(* IEC 61131-3 sources: 2026_Projet_YGO_ExcavatriceDragage/CODE_BACKUP/CODE_20260803_avant_ee4d08b/ACQUISITION, 1 file *)

(* ---- FB_AcquisitionLegacyBridge.st ---- *)
(* ═══════════════════════════════════════════════════════════════
   📡 FB_AcquisitionLegacyBridge — Pont temporaire acquisition historique
   ───────────────────────────────────────────────────────────────
   📄 Docs : DOC/AF_Partie-06_Acquisition_Qualification_IO_v2.0.md §2 ;
            DOC/AF_Partie-13_Fonction_Simulation_v2.0.md
   ⚙️ Pont ST temporaire appelé exclusivement par PRG_02_Acquisition_CFC.xml.
   🎯 Rôle unique : produire l'image matérielle HwIn consommée par le reste
      du programme. Aucune décision métier (SafeStop, mode, commande) ici.
   🔗 Producteur unique de HwIn ; consommateurs = PRG_01_Inputs_LD et suivants.
   ═══════════════════════════════════════════════════════════════ *)

FUNCTION_BLOCK FB_AcquisitionLegacyBridge

VAR_OUTPUT
    HwReal                   : ST_HardwareImage;  (* Image matérielle brute lue sur le terrain *)
    HwSim                    : ST_HardwareImage;  (* Image produite par le banc de simulation *)
    HwIn                     : ST_HardwareImage;  (* Image aiguillée réel/simulé *)
    WinchInputSourceChanged  : BOOL;              (* Pulse 1 cycle sur bascule réel/simulé domaine Winch *)

    // 🆕 Migration PRG_00_Inputs : positions Translation M3 exposées en sortie de programme
    TranslationPosTremie      : BOOL;   (* TRUE = translation en position Trémie *)
    TranslationPosPV          : BOOL;   (* TRUE = translation en zone pré-ralentissement PV *)
    TranslationPosP2          : BOOL;   (* TRUE = translation en position P2 *)
    TranslationPosP1          : BOOL;   (* TRUE = translation en position P1 *)
    TranslationPosMaintenance : BOOL;   (* TRUE = translation en position Maintenance *)

    // 🆕 Migration PRG_00_Inputs : retours variateur M3 filtrés (PT1 T#0MS = recopie legacy)
    M3_StatusWord_Filtered        : UINT;
    M3_ActualFrequencyHz_Filtered : UINT;

    // 🔗 Contrat public : anciennement lus à travers instPosDecoderM3.
    //    Les sorties rendent la migration XML transparente aux consommateurs.
    M3_LimitSwitchFwd          : BOOL;
    M3_LimitSwitchRev          : BOOL;
    M3_SensorWordIncoherent    : BOOL;
    M3_SensorsWord             : BYTE;
END_VAR

VAR
    (* ── Instances de traitement complexes ── *)
    instSimBench             : FB_SimBench;
    instJoystick             : FB_Joystick;
    instEncoderAbsM1         : FB_Encoder_Abs;
    instEncoderScaleM1       : FB_Encoder_Scale;
    instHomingM1             : FB_Encoder_Homing;
    instEncoderAbsM2         : FB_Encoder_Abs;
    instEncoderScaleM2       : FB_Encoder_Scale;
    instHomingM2             : FB_Encoder_Homing;
    instPosDecoderM3         : FB_Translation_PositionDecoder;

    (* ── Filtrage des retours variateur M3 (migration PRG_00_Inputs) ── *)
    instCycleTimeAcq            : FB_CycleTime;
    instFilterM3StatusWord      : FB_Filter_PT1;
    instFilterM3ActualFreqHz      : FB_Filter_PT1;

    (* ── Mémoire de la source Winch (front bascule réel/simulé) ── *)
    WinchInputSourceSimulated            : BOOL;
    PreviousWinchInputSourceSimulated    : BOOL;
    WinchInputSourceInitialized          : BOOL;
END_VAR

// === IMPLEMENTATION ===

// ─── §0 MATÉRIEL ──► HwReal (Acquisition brute unique) ─────────────────────────

// Winch M1 / M2 et codeurs
HwReal.Winch.M1_ContactorsReleased_DI := M1_ContactorsReleased_DI;
HwReal.Winch.M1_ThermalOk_DI          := M1_ThermalOk_DI;
HwReal.Winch.M1_BrakeIsOpen_DI        := M1_BrakeIsOpen_DI;

HwReal.Winch.M2_ContactorsReleased_DI := M2_ContactorsReleased_DI;
HwReal.Winch.M2_ThermalOk_DI          := M2_ThermalOk_DI;
HwReal.Winch.M2_BrakeIsOpen_DI        := M2_BrakeIsOpen_DI;

HwReal.Winch.M1M2_TopPositionFree_DI  := M1M2_TopPositionFree_DI;
HwReal.Winch.M2_TensionedCable_DI     := M2_TensionedCable_DI;

HwReal.Winch.COD1_PosValue            := COD1_PosValue;
HwReal.Winch.COD1_Alarms              := COD1_Alarms;
HwReal.Winch.COD1_Warnings            := COD1_Warnings;
HwReal.Winch.COD1_DeviceState         := COD1_CODEUR.GetDeviceState();

HwReal.Winch.COD2_PosValue            := COD2_PosValue;
HwReal.Winch.COD2_Alarms              := COD2_Alarms;
HwReal.Winch.COD2_Warnings            := COD2_Warnings;
HwReal.Winch.COD2_DeviceState         := COD2_CODEUR.GetDeviceState();

// Translation M3 et variateur AC600
HwReal.Translation.M3_PosTremie_DI      := M3_PosTremie_DI;
HwReal.Translation.M3_PosPV_DI          := M3_PosPV_DI;
HwReal.Translation.M3_PosP2_DI          := M3_PosP2_DI;
HwReal.Translation.M3_PosP1_DI          := M3_PosP1_DI;
HwReal.Translation.M3_PosMaintenance_DI := M3_PosMaintenance_DI;
HwReal.Translation.M3_BrakeIsOpen_DI    := M3_BrakeIsOpen_DI;
HwReal.Translation.M3_ThermalFeedback_DI:= M3_ThermalFeedback_DI; // 🆕 T96 — diagnostic seul (voie déjà mappée CODESYS, jamais lue jusqu'ici)
HwReal.Translation.M3_StatusWord        := M3_StatusWord;
HwReal.Translation.M3_ActualFrequencyHz := M3_ActualFrequencyHz;
HwReal.Translation.AC600_DeviceState    := AC600_ECAT_Drive.GetDeviceState();

// Opérateur / Joystick / bus CANopen
HwReal.Operator.JoyXRaw_ANA1      := JoyXRaw_ANA1;
HwReal.Operator.JoyYRaw_ANA2      := JoyYRaw_ANA2;
HwReal.Operator.JoyBtnRaw         := JoyBtnRaw;
HwReal.Operator.CanBusState       := CANbus.GetBusState();
HwReal.Operator.JOY1_DeviceState  := JOY1_JOYSTICK_MCB560_CO4201A.GetDeviceState();

// Sécurités / Communs Machine
HwReal.Machine.PowerContactorEngaged_DI   := PowerContactorEngaged_DI;
HwReal.Machine.EmergencyChainClosed_DI    := EmergencyChainClosed_DI;
HwReal.Machine.PhaseRotationOk_DI         := PhaseRotationOk_DI;
HwReal.Machine.BrakeThermalOk_DI          := BrakeThermalOk_DI;
HwReal.Machine.M1_M2_KoboldContactFond_DI := M1_M2_KoboldContactFond_DI;
HwReal.Machine.HydraulicThermalOk_DI      := HydraulicThermalOk_DI;

// ─── §0bis HwReal / SimBench ──► HwIn (Aiguillage simulation par domaine) ──────

instSimBench(
    Enable                   := GVL_Simulation.SimulationModeActive,
    M1_RelayFwd              := GVL_Global.M1RelayFwd,
    M1_RelayRev              := GVL_Global.M1RelayRev,
    M1_SpeedContactor_1      := GVL_Global.M1SpeedContactor1,
    M1_SpeedContactor_2      := GVL_Global.M1SpeedContactor2,
    M1_SpeedContactor_3      := GVL_Global.M1SpeedContactor3,
    M1_SpeedContactor_4      := GVL_Global.M1SpeedContactor4,
    M1_SpeedRefPct           := PRG_TREUILS_CFC.M1_SpeedRef_Active,
    M1_PresetTriggerCmd      := PRG_02_Encoders.instEncoderAbsM1.PresetTriggerCmd,
    M1_PresetValueOut        := PRG_02_Encoders.instEncoderAbsM1.PresetValueOut,
    M1_BrakeCmd              := GVL_Global.M1BrakeCmd,
    M2_RelayFwd              := GVL_Global.M2RelayFwd,
    M2_RelayRev              := GVL_Global.M2RelayRev,
    M2_SpeedContactor_1      := GVL_Global.M2SpeedContactor1,
    M2_SpeedContactor_2      := GVL_Global.M2SpeedContactor2,
    M2_SpeedContactor_3      := GVL_Global.M2SpeedContactor3,
    M2_SpeedContactor_4      := GVL_Global.M2SpeedContactor4,
    M2_SpeedRefPct           := PRG_TREUILS_CFC.M2_SpeedRef_Active,
    M2_PresetTriggerCmd      := PRG_02_Encoders.instEncoderAbsM2.PresetTriggerCmd,
    M2_PresetValueOut        := PRG_02_Encoders.instEncoderAbsM2.PresetValueOut,
    M2_BrakeCmd              := GVL_Global.M2BrakeCmd,
    M3_Direction             := PRG_TRANSLATION_CFC.M3_Direction_Active,
    M3_SpeedRefPct           := PRG_TRANSLATION_CFC.M3_SpeedRef_Active,
    M3_BrakeCmd              := GVL_Global.TranslationBrakeCmd,
    M3_TargetNum             := GVL_IHM.TranslationM3.Cmd.SelTarget,
    PowerKeepAlive_A         := PRG_10_Outputs_LD.PowerKeepAlive_A_RQ,
    PowerKeepAlive_B         := PRG_10_Outputs_LD.PowerKeepAlive_B_RQ,
    EmergencyArming_RQ       := PRG_10_Outputs_LD.EmergencyArming_RQ,
    SimEncoderSpeedFactor    := GVL_Simulation.SimEncoderSpeedFactor,
    SimSyncDeviationInjectM1 := GVL_Simulation.SimSyncDeviationInjectM1,
    SimSyncDeviationInjectM2 := GVL_Simulation.SimSyncDeviationInjectM2,
    SimSyncDeviationOffset_M := GVL_Simulation.SimSyncDeviationOffset_M,
    SimM3SensorsWordActive   := GVL_Simulation.SimM3SensorsWordActive,
    SimM3SensorsWord         := GVL_Simulation.SimM3SensorsWord,
    SimJoystickRawX          := GVL_Simulation.SimJoystickRawX,
    SimJoystickRawY          := GVL_Simulation.SimJoystickRawY,
    SimJoystickRawButton     := GVL_Simulation.SimJoystickRawButton,
    SimKoboldContactValue    := GVL_Simulation.SimKoboldContactValue,
    BtnEmergencyStop         := GVL_IHM.Modes.Cmd.BtnEmergencyCutOff,
    HwReal                   := HwReal,
    RawPosM1                 := _SimEncoderRawPosM1,
    RawPosM2                 := _SimEncoderRawPosM2
);

// 🧪 Image du banc exposée pour lecture côte à côte ; aucune logique métier ne lit HwSim.
HwSim.Winch       := instSimBench.Winch;
HwSim.Translation := instSimBench.Translation;
HwSim.Operator    := instSimBench.Operator;
HwSim.Machine     := instSimBench.Machine;

// 🔄 Source Winch atomique + pulse générique. Au boot, la source initiale est mémorisée sans faux pulse.
WinchInputSourceSimulated := GVL_Simulation.SimulationModeActive AND GVL_Simulation.SimWinchActive;
IF NOT WinchInputSourceInitialized THEN
    PreviousWinchInputSourceSimulated := WinchInputSourceSimulated;
    WinchInputSourceInitialized := TRUE;
    WinchInputSourceChanged := FALSE;
ELSE
    WinchInputSourceChanged := (WinchInputSourceSimulated <> PreviousWinchInputSourceSimulated);
    PreviousWinchInputSourceSimulated := WinchInputSourceSimulated;
END_IF;

// Aiguillage domaine par domaine (réel si simulateur inactif pour ce domaine).
IF WinchInputSourceSimulated
    THEN HwIn.Winch := instSimBench.Winch;             ELSE HwIn.Winch := HwReal.Winch;             END_IF;
IF GVL_Simulation.SimulationModeActive AND GVL_Simulation.SimTranslationActive
    THEN HwIn.Translation := instSimBench.Translation; ELSE HwIn.Translation := HwReal.Translation; END_IF;
IF GVL_Simulation.SimulationModeActive AND GVL_Simulation.SimOperatorActive
    THEN HwIn.Operator := instSimBench.Operator;       ELSE HwIn.Operator := HwReal.Operator;       END_IF;
IF GVL_Simulation.SimulationModeActive AND GVL_Simulation.SimMachineActive
    THEN HwIn.Machine := instSimBench.Machine;         ELSE HwIn.Machine := HwReal.Machine;         END_IF;

// ─── §1 TRAITEMENT DES ENTRÉES COMPLEXES (depuis HwIn) ───────────────────────

// 🕹️ Joystick : acquisition + homme-mort + mise à l'échelle
instJoystick(
    Enable                    := TRUE,
    Reset                     := PRG_SUPERVISION_CFC.FaultMachineReset_IHM,
    PowerContactorEngaged     := HwIn.Machine.PowerContactorEngaged_DI,
    Mode                      := PRG_MODES_CFC.Auth.Mode,
    BenneBusy                 := PRG_TREUILS_CFC.instBucket.Busy,
    PreserveArmingAfterBucket := PRG_TREUILS_CFC.instExtractionSequence.Busy
                                 AND (PRG_TREUILS_CFC.instExtractionSequence.ExtractionState = E_ExtractionSequenceState.CLOSING_BUCKET),
    BusCanOpenOP              := PRG_01_Diagnostics.instDiagCanOpen.DeviceCanOpenMaster,
    JoystickOP                := PRG_01_Diagnostics.instDiagCanOpen.DeviceJoystick,
    RawX                      := HwIn.Operator.JoyXRaw_ANA1,
    RawY                      := HwIn.Operator.JoyYRaw_ANA2,
    RawButton                 := HwIn.Operator.JoyBtnRaw,
    BtnCalibrate              := GVL_IHM.JOY1Joystick.Cmd.BtnCalibrate,
    InvertX                   := _JoystickInvertX,
    InvertY                   := _JoystickInvertY,
    Deadband                  := _JoystickDeadband_Pct,
    FilterTime                := _JoystickFilterTime,
    DeadmanRearmTimeout       := T#10S,
    NeutralHoldTime           := T#500MS,
    NeutralXMem               := _JoystickNeutralX,
    NeutralYMem               := _JoystickNeutralY
);

// 🧲 Codeurs M1 : Abs → Homing → Scale
instEncoderAbsM1(
    Enable              := TRUE,
    Reset               := PRG_SUPERVISION_CFC.FaultMachineReset_IHM,
    PowerContactorEngaged     := HwIn.Machine.PowerContactorEngaged_DI,
    Mode                := PRG_MODES_CFC.Auth.Mode,
    RawPosIn            := HwIn.Winch.COD1_PosValue,
    AlarmsIn            := HwIn.Winch.COD1_Alarms,
    WarningsIn          := HwIn.Winch.COD1_Warnings,
    SlaveOperational    := PRG_01_Diagnostics.instDiagEthercat.DeviceEncoderM1.Operational,
    PresetRequest       := instHomingM1.PresetRequest,
    PresetValue         := instHomingM1.PresetValue
);

instHomingM1(
    Enable               := TRUE,
    Reset                := PRG_SUPERVISION_CFC.FaultMachineReset_IHM,
    PowerContactorEngaged      := HwIn.Machine.PowerContactorEngaged_DI,
    Mode                 := PRG_MODES_CFC.Auth.Mode,
    Home                 := GVL_IHM.M1TreuilRetenue.Cmd.BtnHome OR GVL_IHM.M1TreuilRetenue.Cmd.BtnHomingAtZero,
    UnitaryMode          := (PRG_MODES_CFC.Auth.Mode = E_Mode.MAINT_N2)
                            AND (PRG_MODES_CFC.Auth.JoystickWinchSelectArbitrated <> 3),
    WinchSelected        := (PRG_MODES_CFC.Auth.JoystickWinchSelectArbitrated = 1),
    CfgHomingTargetM        := _WinchM1CfgPersist.CfgHomingTarget_M,
    BtnConfirmCoherence     := GVL_IHM.M1TreuilRetenue.Cmd.BtnConfirmCoherence,
    TopPositionSensor    := HwIn.Winch.M1M2_TopPositionFree_DI,
    CfgTopSensorPosM   := SEL(GVL_IHM.M1TreuilRetenue.Cmd.BtnHomingAtZero, _WinchM1CfgPersist.CfgTopSensorPos_M, 0.0),
    FwdRevSpeedFeedbackOff := HwIn.Winch.M1_ContactorsReleased_DI,
    BrakeFeedback        := HwIn.Winch.M1_BrakeIsOpen_DI,
    RawPos               := instEncoderAbsM1.RawPos,
    EncoderAvailable     := instEncoderAbsM1.EncoderAvailable,
    PresetAck            := instEncoderAbsM1.PresetAck,
    PresetNak            := instEncoderAbsM1.PresetNak,
    PointsPerRev         := 8192,
    MultiTurnRevsMax     := 4096,
    CableM_PerRev        := 2.0,
    BypassGlobal         := GVL_IHM.M1TreuilRetenue.Bypass.Global,
    Calib                := _CalibM1
);

instEncoderScaleM1(
    RawPos          := instEncoderAbsM1.RawPos,
    HomingRefRaw    := instHomingM1.HomingRefRaw,
    CableM_PerRev   := 2.0,
    PointsPerRev    := 8192
);

// 🧲 Codeurs M2 : Abs → Homing → Scale
instEncoderAbsM2(
    Enable              := TRUE,
    Reset               := PRG_SUPERVISION_CFC.FaultMachineReset_IHM,
    PowerContactorEngaged     := HwIn.Machine.PowerContactorEngaged_DI,
    Mode                := PRG_MODES_CFC.Auth.Mode,
    RawPosIn            := HwIn.Winch.COD2_PosValue,
    AlarmsIn            := HwIn.Winch.COD2_Alarms,
    WarningsIn          := HwIn.Winch.COD2_Warnings,
    SlaveOperational    := PRG_01_Diagnostics.instDiagEthercat.DeviceEncoderM2.Operational,
    PresetRequest       := instHomingM2.PresetRequest,
    PresetValue         := instHomingM2.PresetValue
);

instHomingM2(
    Enable               := TRUE,
    Reset                := PRG_SUPERVISION_CFC.FaultMachineReset_IHM,
    PowerContactorEngaged      := HwIn.Machine.PowerContactorEngaged_DI,
    Mode                 := PRG_MODES_CFC.Auth.Mode,
    Home                 := GVL_IHM.M2TreuilBenne.Cmd.BtnHome OR GVL_IHM.M2TreuilBenne.Cmd.BtnHomingAtZero,
    UnitaryMode          := (PRG_MODES_CFC.Auth.Mode = E_Mode.MAINT_N2)
                            AND (PRG_MODES_CFC.Auth.JoystickWinchSelectArbitrated <> 3),
    WinchSelected        := (PRG_MODES_CFC.Auth.JoystickWinchSelectArbitrated = 2),
    CfgHomingTargetM        := _WinchM2CfgPersist.CfgHomingTarget_M,
    BtnConfirmCoherence     := GVL_IHM.M2TreuilBenne.Cmd.BtnConfirmCoherence,
    TopPositionSensor    := HwIn.Winch.M1M2_TopPositionFree_DI,
    CfgTopSensorPosM   := SEL(GVL_IHM.M2TreuilBenne.Cmd.BtnHomingAtZero, _WinchM2CfgPersist.CfgTopSensorPos_M, 0.0),
    FwdRevSpeedFeedbackOff := HwIn.Winch.M2_ContactorsReleased_DI,
    BrakeFeedback        := HwIn.Winch.M2_BrakeIsOpen_DI,
    RawPos               := instEncoderAbsM2.RawPos,
    EncoderAvailable     := instEncoderAbsM2.EncoderAvailable,
    PresetAck            := instEncoderAbsM2.PresetAck,
    PresetNak            := instEncoderAbsM2.PresetNak,
    PointsPerRev         := 8192,
    MultiTurnRevsMax     := 4096,
    CableM_PerRev        := 2.0,
    BypassGlobal         := GVL_IHM.M2TreuilBenne.Bypass.Global,
    Calib                := _CalibM2
);

instEncoderScaleM2(
    RawPos          := instEncoderAbsM2.RawPos,
    HomingRefRaw    := instHomingM2.HomingRefRaw,
    CableM_PerRev   := 2.0,
    PointsPerRev    := 8192
);

// ↔️ Translation M3 : décodage du mot de capteurs de position
instPosDecoderM3(
    SensorTremie      := HwIn.Translation.M3_PosTremie_DI,
    SensorPV          := HwIn.Translation.M3_PosPV_DI,
    SensorP2          := HwIn.Translation.M3_PosP2_DI,
    SensorP1          := HwIn.Translation.M3_PosP1_DI,
    SensorMaintenance := HwIn.Translation.M3_PosMaintenance_DI
);

// 🆕 Exposition des positions Translation M3 pour les consommateurs legacy
TranslationPosTremie      := instPosDecoderM3.TranslationPosTremie;
TranslationPosPV          := instPosDecoderM3.TranslationPosPV;
TranslationPosP2          := instPosDecoderM3.TranslationPosP2;
TranslationPosP1          := instPosDecoderM3.TranslationPosP1;
TranslationPosMaintenance := instPosDecoderM3.TranslationPosMaintenance;
M3_LimitSwitchFwd       := instPosDecoderM3.LimitSwitchFwd;
M3_LimitSwitchRev       := instPosDecoderM3.LimitSwitchRev;
M3_SensorWordIncoherent := instPosDecoderM3.Incoherent;
M3_SensorsWord          := instPosDecoderM3.SensorsWord;

// 🆕 Filtrage PT1 (T#0MS = pass-through) des retours variateur M3 — cohérent avec le legacy
instCycleTimeAcq(DefaultValueS := 0.010);

instFilterM3StatusWord(
    ValueIn    := UINT_TO_REAL(WORD_TO_UINT(HwIn.Translation.M3_StatusWord)),
    TimeConst  := T#0MS,
    CycleTimeS := instCycleTimeAcq.CycleTimeS
);
M3_StatusWord_Filtered := REAL_TO_UINT(instFilterM3StatusWord.ValueOut);

instFilterM3ActualFreqHz(
    ValueIn    := UINT_TO_REAL(HwIn.Translation.M3_ActualFrequencyHz),
    TimeConst  := T#0MS,
    CycleTimeS := instCycleTimeAcq.CycleTimeS
);
M3_ActualFrequencyHz_Filtered := REAL_TO_UINT(instFilterM3ActualFreqHz.ValueOut);
